(* IEC 61131-3 sources: SortJet_MasterSPS_Aufbau.fbsproj/09_Station/Stationen/Anlegetisch[201,205]/0_Unterbausteine, 2 files *)

(* ---- ZylinderPneumatik_Anschlag_FB_V01_00_00.fb.st ---- *)
(* METADATA
{
	"v3Meta": {
		"objectGuid": "73b344ea-77d6-4df9-8490-b74a4c5cebf9"
	}
}
*)
FUNCTION_BLOCK ZylinderPneumatik_Anschlag_FB_V01_00_00
VAR_INPUT

  // EINGAENGE
  in_bStatusZylinderAusgefahren : BOOL;
  in_bStatusZylinderEingefahren : BOOL;

  // BOOLEAN
  bpReset                       : BOOL;
  bpAktivieren                  : BOOL;
  bpFreigabe                    : BOOL; // FREIGABE Pneumatik: ohne Freigabe Ventile aus, Bewegung pausiert (Startbefehl bleibt erhalten)
  bpStartAusfahren              : BOOL;
  bpStartEinfahren              : BOOL;

  // OPTIONEN
  bpAbfrageAusgefahrenVorhanden : BOOL := TRUE;   // Endlagensensor ausgefahren vorhanden, sonst gilt die Endlage nach tpBewegungszeit
  bpAbfrageEingefahrenVorhanden : BOOL := TRUE;   // Endlagensensor eingefahren vorhanden, sonst gilt die Endlage nach tpBewegungszeit
  tpBewegungszeit               : TIME := T#800MS; // Bewegungszeit je Richtung ohne Endlagensensor

END_VAR
VAR_OUTPUT
  // AUSGAENGE
  out_bZylinderAusfahren        : BOOL;
  out_bZylinderEinfahren        : BOOL;

  // BOOLEAN
  bpFehler                      : BOOL;
  bpDone                        : BOOL;

  // WORD
  wpFehlerNr                    : Fehlerkonstanten_EN;

  // ENUM
  epStatusZylinder : PneumatikZylinderStatus_EN;

END_VAR
VAR

  // STEPS
  steplAusfahren   : Steps_TE;
  steplEinfahren   : Steps_TE;

  // TIMER
  tonZylinderEingefahren     : TON; // EINSCHALTVERZOEGERUNG: Warten bis der Zylinder eingefahren wurde. Sonst wird ein Fehlerausgegeben
  tonZylinderAusgefahren     : TON; // EINSCHALTVERZOEGERUNG: Warten bis der Zylinder ausgefahren wurde. Sonst wird ein Fehlerausgegeben
  tonlBewegungszeitEinfahren : TON; // Bewegungszeit ohne Endlagensensor eingefahren
  tonlBewegungszeitAusfahren : TON; // Bewegungszeit ohne Endlagensensor ausgefahren

END_VAR

VAR CONSTANT

  // TIME
  cZEITLICHE_UEBERWACHUNG_BEWEGUNG_ZYLINDER : TIME := T#15s;

END_VAR
//-------------------------------------------------------------------------------------------------
// BAUSTEIN: RESET / DEAKTIVIERT
//-------------------------------------------------------------------------------------------------
(* Hinweis:
   - Reset oder deaktiviert: Ausgaenge aus, Ketten und Timer zuruecksetzen, Done und Fehler loeschen
   - Der Baustein setzt bpReset selbst zurueck, der Aufrufer wartet nicht auf Done
   - Ein deaktivierter Zylinder meldet kein Done; der Aufrufer verknuepft das Warten auf Done
     mit der Aktivierung aus der MK (z.B. Zylinder.bpDone OR NOT stStationsAufbau.bX)
*)
IF ( bpReset OR NOT bpAktivieren ) THEN

  out_bZylinderAusfahren := FALSE;
  out_bZylinderEinfahren := FALSE;

  bpStartAusfahren := FALSE;
  bpStartEinfahren := FALSE;

  steplAusfahren := STEP_0_E;
  steplEinfahren := STEP_0_E;

  tonZylinderAusgefahren( IN := FALSE );
  tonZylinderEingefahren( IN := FALSE );
  tonlBewegungszeitAusfahren( IN := FALSE );
  tonlBewegungszeitEinfahren( IN := FALSE );

  bpDone     := FALSE;
  bpFehler   := FALSE;
  wpFehlerNr := cMELDUNG_NULL;

  bpReset := FALSE;

  RETURN;

END_IF

//-------------------------------------------------------------------------------------------------
// BAUSTEIN: AKTIONEN
//-------------------------------------------------------------------------------------------------
(* Hinweis Freigabe Pneumatik:
   - Ohne Freigabe: Ventile aus, Ketten und Ueberwachungszeiten zuruecksetzen (kein Timeout-Fehler)
   - Der Startbefehl bleibt erhalten: kommt die Freigabe zurueck, wird die Bewegung neu gestartet
*)
IF NOT bpFreigabe THEN
  out_bZylinderAusfahren := FALSE;
  out_bZylinderEinfahren := FALSE;
  steplAusfahren := STEP_0_E;
  steplEinfahren := STEP_0_E;
  tonZylinderAusgefahren( IN := FALSE );
  tonZylinderEingefahren( IN := FALSE );
  tonlBewegungszeitAusfahren( IN := FALSE );
  tonlBewegungszeitEinfahren( IN := FALSE );
  bpDone := FALSE;
ELSE
  Ausfahren();
  Einfahren();
END_IF

//-------------------------------------------------------------------------------------------------
// STATUS DES ZYLINDERS
//-------------------------------------------------------------------------------------------------
(* Hinweis:
   - Status aus der Sensorik, soweit Endlagensensoren vorhanden sind
   - Ohne Sensor bleibt der Status, den die Schrittketten nach der Bewegungszeit setzen
*)
IF ( bpAbfrageAusgefahrenVorhanden AND bpAbfrageEingefahrenVorhanden ) THEN

  IF (      in_bStatusZylinderAusgefahren
       AND NOT in_bStatusZylinderEingefahren )
  THEN
    epStatusZylinder := eZylinderAusgefahren;
  ELSIF(    in_bStatusZylinderEingefahren
         AND NOT in_bStatusZylinderAusgefahren )
  THEN
    epStatusZylinder := eZylinderEingefahren;
  ELSE
    epStatusZylinder := eZylinderUndefiniert;
  END_IF

ELSIF ( bpAbfrageAusgefahrenVorhanden ) THEN

  IF ( in_bStatusZylinderAusgefahren ) THEN
    epStatusZylinder := eZylinderAusgefahren;
  ELSIF ( epStatusZylinder = eZylinderAusgefahren ) THEN
    epStatusZylinder := eZylinderUndefiniert;
  END_IF

ELSIF ( bpAbfrageEingefahrenVorhanden ) THEN

  IF ( in_bStatusZylinderEingefahren ) THEN
    epStatusZylinder := eZylinderEingefahren;
  ELSIF ( epStatusZylinder = eZylinderEingefahren ) THEN
    epStatusZylinder := eZylinderUndefiniert;
  END_IF

END_IF
END_FUNCTION_BLOCK

(* ---- ZylinderPneumatik_Riemen_FB_V01_00_00.fb.st ---- *)
(* METADATA
{
	"v3Meta": {
		"objectGuid": "4bd964be-8117-422d-b97f-60e1c4b0ab77"
	}
}
*)
FUNCTION_BLOCK ZylinderPneumatik_Riemen_FB_V01_00_00
VAR_INPUT
  // HARDWARE EINGAENGE
  in_bStatusZylinderAusgefahren : BOOL; // STATUS: Sensor meldt ausgfahren
  in_bStatusZylinderEingefahren : BOOL; // STATUS: Sensor meldt eingefahren

  // BOOLEAN
  bpAktivieren     : BOOL; // AKTIVIERUNG: stStationsAufbau.bHubrahmen
  bpFreigabe       : BOOL; // FREIGABE Pneumatik: ohne Freigabe Ventil aus (Feder faehrt zurueck), Bewegung pausiert (Startbefehl bleibt erhalten)
  bpStartAusfahren : BOOL; // BETRIEBTYP: Zylinder wird ausgefahren
  bpStartEinfahren : BOOL; // BETRIEBTYP: Zylinder wird eingefahren
  bpReset          : BOOL; // BETRIEBTYP: Zylinderbaustein wird zurueckgesetzt

  // OPTIONEN
  bpAbfrageAusgefahrenVorhanden : BOOL := TRUE;   // Endlagensensor ausgefahren vorhanden, sonst gilt die Endlage nach tpBewegungszeit
  bpAbfrageEingefahrenVorhanden : BOOL := TRUE;   // Endlagensensor eingefahren vorhanden, sonst gilt die Endlage nach tpBewegungszeit
  tpBewegungszeit               : TIME := T#800MS; // Bewegungszeit je Richtung ohne Endlagensensor

END_VAR
VAR_OUTPUT
  // HARDWARE AUSGAENGE
  out_bZylinderAusfahren : BOOL; // AUSGANG: (in Glasflussrichtung) Signal zum Ausfahren  [Federrueckstell- Ventiel]

  // BOOLEAN
  bpFehler   : BOOL;
  bpDone     : BOOL;

  // WORD
  wpFehlerNr : Fehlerkonstanten_EN;

  // ENUM
  epStatusZylinder : PneumatikZylinderStatus_EN;

END_VAR
VAR
  // STEPS
  steplAusfahren   : Steps_TE;
  steplEinfahren   : Steps_TE;

  // TIMER
  tonlZylinderEingefahren    : TON; // EINSCHALTVERZOEGERUNG: Warten bis der Zylinder eingefahren wurde. Sonst wird ein Fehlerausgegeben
  tonlZylinderAusgefahren    : TON; // EINSCHALTVERZOEGERUNG: Warten bis der Zylinder ausgefahren wurde. Sonst wird ein Fehlerausgegeben
  tonlBewegungszeitEinfahren : TON; // Bewegungszeit ohne Endlagensensor eingefahren
  tonlBewegungszeitAusfahren : TON; // Bewegungszeit ohne Endlagensensor ausgefahren

END_VAR
VAR CONSTANT

  // TIME
  cZEITLICHE_UEBERWACHUNG_BEWEGUNG_ZYLINDER : TIME := T#5s;

END_VAR
(* Hinweis:
   - Es handelt sich bei diesem Baustein um eine Ansteuerung fuer ein Federrueckstell- Ventiel
     => Der Ausgang bleibt nach dem Ausfahren gesetzt, Einfahren nimmt ihn zurueck
*)

//-------------------------------------------------------------------------------------------------
// BAUSTEIN: RESET / DEAKTIVIERT
//-------------------------------------------------------------------------------------------------
(* Hinweis:
   - Reset oder deaktiviert: Ausgang aus, Ketten und Timer zuruecksetzen, Done und Fehler loeschen
   - Der Baustein setzt bpReset selbst zurueck, der Aufrufer wartet nicht auf Done
   - Ein deaktivierter Zylinder meldet kein Done; der Aufrufer verknuepft das Warten auf Done
     mit der Aktivierung aus der MK (z.B. Zylinder.bpDone OR NOT stStationsAufbau.bX)
*)
IF ( bpReset OR NOT bpAktivieren ) THEN

  out_bZylinderAusfahren := FALSE;

  bpStartAusfahren := FALSE;
  bpStartEinfahren := FALSE;

  steplAusfahren := STEP_0_E;
  steplEinfahren := STEP_0_E;

  tonlZylinderAusgefahren( IN := FALSE );
  tonlZylinderEingefahren( IN := FALSE );
  tonlBewegungszeitAusfahren( IN := FALSE );
  tonlBewegungszeitEinfahren( IN := FALSE );

  bpDone     := FALSE;
  bpFehler   := FALSE;
  wpFehlerNr := cMELDUNG_NULL;

  bpReset := FALSE;

  RETURN;

END_IF

//-------------------------------------------------------------------------------------------------
// BAUSTEIN: AKTIONEN
//-------------------------------------------------------------------------------------------------
(* Hinweis Freigabe Pneumatik:
   - Ohne Freigabe: Ventil aus, Ketten und Ueberwachungszeiten zuruecksetzen (kein Timeout-Fehler)
   - Der Startbefehl bleibt erhalten: kommt die Freigabe zurueck, wird die Bewegung neu gestartet
*)
IF NOT bpFreigabe THEN
  out_bZylinderAusfahren := FALSE;
  steplAusfahren := STEP_0_E;
  steplEinfahren := STEP_0_E;
  tonlZylinderAusgefahren( IN := FALSE );
  tonlZylinderEingefahren( IN := FALSE );
  tonlBewegungszeitAusfahren( IN := FALSE );
  tonlBewegungszeitEinfahren( IN := FALSE );
  bpDone := FALSE;
ELSE
  Ausfahren();
  Einfahren();
END_IF

//-------------------------------------------------------------------------------------------------
// STATUS DES ZYLINDERS
//-------------------------------------------------------------------------------------------------
(* Hinweis:
   - Status aus der Sensorik, soweit Endlagensensoren vorhanden sind
   - Ohne Sensor bleibt der Status, den die Schrittketten nach der Bewegungszeit setzen
*)
IF ( bpAbfrageAusgefahrenVorhanden AND bpAbfrageEingefahrenVorhanden ) THEN

  IF (      in_bStatusZylinderAusgefahren
       AND NOT in_bStatusZylinderEingefahren )
  THEN
    epStatusZylinder := eZylinderAusgefahren;
  ELSIF(    in_bStatusZylinderEingefahren
         AND NOT in_bStatusZylinderAusgefahren )
  THEN
    epStatusZylinder := eZylinderEingefahren;
  ELSE
    epStatusZylinder := eZylinderUndefiniert;
  END_IF

ELSIF ( bpAbfrageAusgefahrenVorhanden ) THEN

  IF ( in_bStatusZylinderAusgefahren ) THEN
    epStatusZylinder := eZylinderAusgefahren;
  ELSIF ( epStatusZylinder = eZylinderAusgefahren ) THEN
    epStatusZylinder := eZylinderUndefiniert;
  END_IF

ELSIF ( bpAbfrageEingefahrenVorhanden ) THEN

  IF ( in_bStatusZylinderEingefahren ) THEN
    epStatusZylinder := eZylinderEingefahren;
  ELSIF ( epStatusZylinder = eZylinderEingefahren ) THEN
    epStatusZylinder := eZylinderUndefiniert;
  END_IF

END_IF
END_FUNCTION_BLOCK
